// TIA Portal project "071_db_1200_300" (V21)

(* hardware
DEVICE "PLC_1200"  S7-1200 Station
   slot 0: "Rack_0"  S7-1200 Rack  Rack  V1.0
   slot 1: "PLC_1200"  CPU 1214C DC/DC/DC  6ES7 214-1AG40-0XB0  V4.7
DEVICE "PLC_300"  S7-300 station
   slot 0: "Rail_0"  Rail  6ES7 390-1***0-0AA0
   slot 2: "PLC_300"  CPU 315-2 PN/DP  6ES7 315-2EH14-0AB0  V3.2
      slot 2: "PROFINET interface_1"  PN-IO
         slot 1: "Port_1"  Port
         slot 2: "Port_2"  Port
*)

// ===== PLC "PLC_1200"  CPU 1214C DC/DC/DC =====

TYPE "UDT_12"
   STRUCT
      "a" : Int := 3;
      "b" : Real;
      c : Array[0..1] of Bool;
   END_STRUCT;
END_TYPE

DATA_BLOCK "DB_12Opt"   // DB1
{ S7_Optimized_Access := 'TRUE' }
   VAR
      x : Bool;
      i : Int := 12;
      d : DInt;
      r : Real;
      lr : LReal;
      t : Time;
      dtl : DTL;
      s : String[10] := 'S7-1200';
      ws : WString;
      a2 : Array[0..1, 0..2] of Int;
      st : Struct
         p : Word;
         q : Array[1..3] of Byte;
      END_STRUCT;
      u : "UDT_12";
      au : Array[0..1] of "UDT_12";
      tm : IEC_TIMER;
   END_VAR
   VAR RETAIN
      rr : UDInt;
   END_VAR
BEGIN
   a2[1,2] := 7;
   u."b" := 2.5;
   au[1]."a" := 9;
END_DATA_BLOCK

DATA_BLOCK "DB_12Std"   // DB2
{ S7_Optimized_Access := 'FALSE' }
   VAR
      b0 : Bool;
      w : Word;
      i : Int := -4;
      r : Real;
      s : String[6];
      arr : Array[0..3] of Int;
      u : "UDT_12";
   END_VAR
BEGIN
   arr[2] := 22;
END_DATA_BLOCK

DATA_BLOCK "FB_12_DB"   // DB3
{ S7_Optimized_Access := 'TRUE' }
VERSION : 0.1
// stored: InstanceOfName FB_12
"FB_12"
BEGIN
END_DATA_BLOCK

FUNCTION_BLOCK "FB_12"   // FB1, SCL
{ S7_Optimized_Access := 'TRUE' }
VERSION : 0.1
   VAR_INPUT
      en1 : Bool;
      par : "UDT_12";
   END_VAR
   VAR_OUTPUT
      q : Int;
   END_VAR
   VAR
      cnt : Int := 5;
      tmr : TON_TIME;
      edge : R_TRIG;
   END_VAR
BEGIN
   #tmr(IN := #en1, PT := T#1S);
           #q := #cnt;
END_FUNCTION_BLOCK

ORGANIZATION_BLOCK "Main"   // OB1, LAD, ProgramCycle
TITLE = "Main Program Sweep (Cycle)"
{ S7_Optimized_Access := 'TRUE' }
VERSION : 0.1
   VAR_INPUT
      Initial_Call : Bool;   // Initial call of this OB
      Remanence : Bool;   // =True, if remanent data are available
   END_VAR
BEGIN
END_ORGANIZATION_BLOCK

// ===== PLC "PLC_300"  CPU 315-2 PN/DP =====

TYPE "UDT_300"
   STRUCT
      "a" : Int := 3;
      "b" : Real;
      c : Array[0..1] of Bool;
   END_STRUCT;
END_TYPE

DATA_BLOCK "DB_300"   // DB1
{ S7_Optimized_Access := 'FALSE' }
   VAR
      x : Bool;
      i : Int := 30;
      d : DInt;
      r : Real := 1.25;
      t : Time;
      dtv : Date_And_Time;
      s : String[8] := 'S7-300';
      arr : Array[0..3] of Int;
      "m" : Array[0..1, 0..1] of Word;
      st : Struct
         p : Word;
         q : Byte;
      END_STRUCT;
      u : "UDT_300";
   END_VAR
BEGIN
   arr[2] := 22;
   "m"[1,1] := WORD#16#ABCD;
END_DATA_BLOCK

DATA_BLOCK "FB_300_DB"   // DB2
{ S7_Optimized_Access := 'FALSE' }
VERSION : 0.1
// stored: InstanceOfName FB_300
"FB_300"
BEGIN
   cnt := 8;
END_DATA_BLOCK

FUNCTION_BLOCK "FB_300"   // FB1, SCL
{ S7_Optimized_Access := 'FALSE' }
   VAR_INPUT
      en1 : Bool;
   END_VAR
   VAR_OUTPUT
      q : Int;
   END_VAR
   VAR
      cnt : Int := 5;
      u : "UDT_300";
   END_VAR
BEGIN

       #q := #cnt;
END_FUNCTION_BLOCK

ORGANIZATION_BLOCK "Main"   // OB1, LAD
TITLE = "Main Program Sweep (Cycle)"
{ S7_Optimized_Access := 'FALSE' }
VERSION : 0.1
   VAR_TEMP
      OB1_EV_CLASS : Byte;   // Bits 0-3 = 1 (Coming event), Bits 4-7 = 1 (Event class 1)
      OB1_SCAN_1 : Byte;   // 1 (Cold restart scan 1 of OB 1), 3 (Scan 2-n of OB 1)
      OB1_PRIORITY : Byte;   // Priority of OB Execution
      OB1_OB_NUMBR : Byte;   // 1 (Organization block 1, OB1)
      OB1_RESERVED_1 : Byte;   // Reserved for system
      OB1_RESERVED_2 : Byte;   // Reserved for system
      OB1_PREV_CYCLE : Int;   // Cycle time of previous OB1 scan (milliseconds)
      OB1_MIN_CYCLE : Int;   // Minimum cycle time of OB1 (milliseconds)
      OB1_MAX_CYCLE : Int;   // Maximum cycle time of OB1 (milliseconds)
      OB1_DATE_TIME : Date_And_Time;   // Date and time OB1 started
   END_VAR
BEGIN
END_ORGANIZATION_BLOCK